Fanuc KAREL source: KA00084.KL

PROGRAM KA00084
%NOLOCKGROUP
VAR
  SRC: XYZWPREXT
  DST: ARRAY[2] OF SHORT
BEGIN
  SRC.X = 1.0
  DST[1] = SRC
END KA00084
